// TIA Portal V19 export
// export: Created 2026-10-15T09:44:24.355296Z, ExportSetting WithDefaults, DisplayName Totally Integrated Automation Portal, DisplayVersion V19, DisplayName TIA Portal Openness, DisplayVersion V19, DisplayName TIA Portal Version Control Interface, DisplayVersion V19, DisplayName STEP 7 Professional, DisplayVersion V19, DisplayName STEP 7 Safety, DisplayVersion V19, DisplayName WinCC Basic/Comfort/Advanced, DisplayVersion V19, DisplayName WinCC Unified, DisplayVersion V19
FUNCTION "ROLL_PB16" : Void   // FC24, SCL
{ S7_Optimized_Access := 'TRUE' }
VERSION : 0.1
// stored: AutoNumber true, IsIECCheckEnabled false, SetENOAutomatically false, UDAEnableTagReadback false
   VAR_TEMP
      r : Bool;
      a1 : Word;
      a2 : Word;
      activeDataBlock : Int;
      comparisonResults : Array[0..0] of Bool;
   END_VAR
BEGIN

   #r := FALSE;
   #a1 := W#16#0000;
   #a2 := W#16#0000;
   #activeDataBlock := 0;
   // PB16, STEP 5 network 1
   #r := ("ROLL_IO".Input[0, 1] AND "ROLL_State".M[190, 5] AND "ROLL_State".M[190, 6] AND "ROLL_State".M[27, 7]);
   "ROLL_State".M[73, 7] := #r;
   // PB16, STEP 5 network 2
   #r := (("ROLL_State".M[20, 3] OR "ROLL_State".M[20, 5]) AND "ROLL_IO".Input[124, 1] AND "ROLL_IO".Input[124, 4]);
   "ROLL_State".M[74, 2] := #r;
   // PB16, STEP 5 network 3
   #r := (((NOT "ROLL_State".M[190, 5]) AND "ROLL_State".M[190, 6] AND "ROLL_State".M[74, 2]) OR (("ROLL_State".M[70, 2] OR "ROLL_State".M[70, 3]) AND "ROLL_State".M[74, 0]));
   "ROLL_State".M[74, 1] := #r;
   // PB16, STEP 5 network 4
   #r := (("ROLL_State".M[20, 4] OR "ROLL_State".M[20, 5]) AND "ROLL_IO".Input[0, 1] AND "ROLL_State".M[190, 6]);
   "ROLL_State".M[74, 4] := #r;
   // PB16, STEP 5 network 5
   #r := ((NOT "ROLL_IO".Output[113, 3]) AND ("ROLL_IO".Input[123, 6] OR "ROLL_State".M[70, 3] OR "ROLL_State".M[70, 5] OR "ROLL_State".M[70, 6]) AND ("ROLL_State".M[74, 0] OR "ROLL_State".M[74, 4]));
   "ROLL_State".M[74, 5] := #r;
   // PB16, STEP 5 network 6
   #r := ((NOT "ROLL_IO".Input[11, 0]) AND (NOT "ROLL_IO".Input[11, 1]) AND (NOT "ROLL_IO".Input[11, 2]) AND (NOT "ROLL_IO".Input[11, 3]) AND (NOT "ROLL_IO".Input[11, 4]) AND (NOT "ROLL_IO".Input[119, 6]) AND (NOT "ROLL_IO".Input[119, 7]) AND (NOT "ROLL_IO".Input[120, 0]) AND (NOT "ROLL_IO".Input[120, 1]));
   "ROLL_State".M[75, 2] := #r;
   // PB16, STEP 5 network 7
   #r := (("ROLL_State".M[190, 6] AND "ROLL_State".M[23, 1] AND "ROLL_State".M[75, 3]) OR "ROLL_State".M[75, 2]);
   "ROLL_State".M[75, 3] := #r;
   // PB16, STEP 5 network 8
   #r := ((((NOT "ROLL_IO".Input[11, 0]) AND (NOT "ROLL_IO".Input[11, 1]) AND (NOT "ROLL_IO".Input[11, 2]) AND (NOT "ROLL_IO".Input[11, 3]) AND (NOT "ROLL_IO".Input[11, 4]) AND (NOT "ROLL_IO".Input[119, 6]) AND (NOT "ROLL_IO".Input[119, 7]) AND (NOT "ROLL_IO".Input[120, 0]) AND (NOT "ROLL_IO".Input[120, 1]) AND "ROLL_IO".Input[13, 3]) OR "ROLL_State".M[63, 1]) AND ((NOT "ROLL_IO".Input[11, 6]) OR (NOT "ROLL_State".M[75, 3]) OR "ROLL_State".M[75, 2]) AND "ROLL_IO".Input[0, 1] AND "ROLL_IO".Input[12, 5] AND "ROLL_State".M[190, 6] AND "ROLL_State".M[23, 1]);
   "ROLL_State".M[75, 4] := #r;
   // PB16, STEP 5 network 9
   #r := ((((NOT "ROLL_IO".Input[11, 0]) AND (NOT "ROLL_IO".Input[11, 1]) AND (NOT "ROLL_IO".Input[11, 2]) AND (NOT "ROLL_IO".Input[11, 3]) AND (NOT "ROLL_IO".Input[11, 4]) AND (NOT "ROLL_IO".Input[119, 6]) AND (NOT "ROLL_IO".Input[119, 7]) AND (NOT "ROLL_IO".Input[120, 0]) AND (NOT "ROLL_IO".Input[120, 1]) AND "ROLL_IO".Input[13, 3]) OR "ROLL_State".M[63, 1]) AND (((NOT "ROLL_State".M[190, 6]) AND "ROLL_State".M[190, 5] AND "ROLL_State".M[23, 1]) OR "ROLL_State".M[74, 0]) AND "ROLL_IO".Input[0, 1]);
   "ROLL_State".M[75, 5] := #r;
   // PB16, STEP 5 network 10
   #r := (((NOT "ROLL_IO".Input[11, 0]) AND (("ROLL_IO".Input[0, 1] AND "ROLL_State".M[190, 5] AND "ROLL_State".M[23, 1]) OR "ROLL_State".M[74, 0]) AND "ROLL_State".M[63, 1]) OR ("ROLL_IO".Input[0, 1] AND "ROLL_State".M[190, 6] AND "ROLL_State".M[23, 1] AND "ROLL_State".M[75, 2]));
   "ROLL_State".M[75, 6] := #r;
   // PB16, STEP 5 network 11
   #r := ((NOT "ROLL_IO".Input[11, 0]) AND "ROLL_IO".Input[11, 6] AND "ROLL_State".M[190, 5] AND "ROLL_State".M[23, 0]);
   "ROLL_State".M[76, 0] := #r;
   // PB16, STEP 5 network 12
   #r := (((NOT "ROLL_IO".Input[11, 0]) AND "ROLL_State".M[74, 0]) OR ("ROLL_IO".Input[11, 0] AND "ROLL_IO".Input[11, 6] AND "ROLL_State".M[190, 6] AND "ROLL_State".M[23, 0]));
   "ROLL_State".M[76, 1] := #r;
   // PB16, STEP 5 network 13
   #r := (("ROLL_State".M[76, 0] OR "ROLL_State".M[76, 1]) AND "ROLL_IO".Input[0, 1]);
   "ROLL_State".M[76, 2] := #r;
   // PB16, STEP 5 network 14
   #r := ((NOT "ROLL_IO".Input[12, 1]) AND (NOT "ROLL_IO".Input[12, 5]));
   "ROLL_State".M[240, 0] := #r;
   // PB16, STEP 5 network 15
   #r := (("ROLL_State".M[190, 6] AND "ROLL_State".M[23, 0] AND "ROLL_State".M[77, 1]) OR "ROLL_State".M[240, 0]);
   "ROLL_State".M[77, 1] := #r;
   // PB16, STEP 5 network 16
   #r := ((((NOT "ROLL_IO".Input[12, 1]) AND ("ROLL_IO".Input[11, 1] OR "ROLL_IO".Input[11, 2] OR "ROLL_IO".Input[11, 3] OR "ROLL_IO".Input[11, 4] OR "ROLL_IO".Input[119, 6] OR "ROLL_IO".Input[119, 7] OR "ROLL_IO".Input[120, 0] OR "ROLL_IO".Input[120, 1])) OR (NOT "ROLL_IO".Input[12, 7])) AND ((NOT "ROLL_IO".Input[12, 7]) OR (NOT "ROLL_State".M[77, 1]) OR "ROLL_State".M[240, 0]) AND "ROLL_IO".Input[0, 1] AND "ROLL_IO".Input[11, 6] AND "ROLL_State".M[190, 6] AND "ROLL_State".M[23, 0]);
   "ROLL_State".M[77, 2] := #r;
   // PB16, STEP 5 network 17
   #r := (((NOT "ROLL_State".M[6, 0]) AND (NOT "ROLL_State".M[6, 2]) AND ("ROLL_IO".Input[11, 1] OR "ROLL_IO".Input[11, 2] OR "ROLL_IO".Input[11, 3] OR "ROLL_IO".Input[11, 4] OR "ROLL_IO".Input[119, 6] OR "ROLL_IO".Input[119, 7] OR "ROLL_IO".Input[120, 0])) OR "ROLL_IO".Input[11, 4]);
   "ROLL_State".M[76, 4] := #r;
   // PB16, STEP 5 network 18
   #r := ((NOT "ROLL_State".M[190, 5]) AND "ROLL_State".M[190, 6] AND "ROLL_State".M[23, 0] AND "ROLL_State".M[76, 4] AND "ROLL_State".M[77, 2]);
   "ROLL_State".M[76, 5] := #r;
   // PB16, STEP 5 network 19
   #r := ((((NOT "ROLL_State".M[190, 6]) AND "ROLL_State".M[190, 5] AND "ROLL_State".M[23, 0]) OR "ROLL_State".M[74, 0]) AND (("ROLL_IO".Input[124, 2] AND "ROLL_IO".Input[124, 5]) OR "ROLL_State".M[0, 4]) AND "ROLL_IO".Input[11, 0] AND "ROLL_State".M[63, 1]);
   "ROLL_State".M[76, 6] := #r;
   // PB16, STEP 5 network 20
   #r := (((((NOT "ROLL_IO".Input[12, 1]) OR (NOT "ROLL_IO".Input[12, 7])) AND "ROLL_State".M[76, 6]) OR "ROLL_State".M[76, 5]) AND "ROLL_IO".Input[0, 1] AND "ROLL_IO".Input[11, 6]);
   "ROLL_State".M[77, 0] := #r;
   // PB16, STEP 5 network 21
   #r := (((NOT "ROLL_IO".Input[11, 0]) AND (NOT "ROLL_IO".Input[12, 5]) AND "ROLL_State".M[190, 5]) OR ((NOT "ROLL_IO".Input[12, 1]) AND "ROLL_IO".Input[11, 0] AND "ROLL_State".M[190, 6]));
   "ROLL_State".M[240, 0] := #r;
   // PB16, STEP 5 network 22
   #r := ((NOT "ROLL_IO".Input[12, 1]) AND ("ROLL_IO".Input[11, 1] OR "ROLL_IO".Input[11, 2] OR "ROLL_IO".Input[11, 3] OR "ROLL_IO".Input[11, 4] OR "ROLL_IO".Input[119, 6] OR "ROLL_IO".Input[119, 7] OR "ROLL_IO".Input[120, 0]));
   "ROLL_State".M[240, 1] := #r;
   // PB16, STEP 5 network 23
   #r := ((NOT "ROLL_IO".Input[12, 1]) AND "ROLL_IO".Input[11, 0]);
   "ROLL_State".M[240, 2] := #r;
   // PB16, STEP 5 network 24
   #r := ((("ROLL_State".M[240, 1] OR "ROLL_State".M[240, 2]) AND "ROLL_State".M[77, 0]) OR ("ROLL_State".M[240, 0] AND "ROLL_State".M[76, 2]));
   "ROLL_State".M[76, 7] := #r;
   // PB16, STEP 5 network 25
   #r := ((NOT "ROLL_IO".Output[113, 3]) AND (NOT "ROLL_State".M[70, 2]) AND (NOT "ROLL_State".M[70, 3]) AND "ROLL_IO".Input[0, 1] AND "ROLL_IO".Input[11, 0] AND "ROLL_IO".Input[12, 1] AND "ROLL_IO".Input[12, 7] AND "ROLL_IO".Input[124, 5]);
   "ROLL_State".M[77, 3] := #r;
   // PB16, STEP 5 network 26
   #r := ((NOT "ROLL_State".M[77, 6]) AND (((NOT "ROLL_State".M[190, 6]) AND "ROLL_State".M[190, 5] AND "ROLL_State".M[22, 0]) OR "ROLL_State".M[74, 0]) AND "ROLL_IO".Output[113, 2] AND "ROLL_State".M[77, 3]);
   "ROLL_State".M[77, 4] := #r;
   // PB16, STEP 5 network 27
   #r := ((NOT "ROLL_State".M[190, 5]) AND (NOT "ROLL_State".M[77, 4]) AND "ROLL_State".M[190, 6] AND "ROLL_State".M[22, 0] AND "ROLL_State".M[77, 3]);
   "ROLL_State".M[77, 6] := #r;
   // PB16, STEP 5 network 28
   #r := ((NOT "ROLL_IO".Input[124, 5]) AND (NOT "ROLL_State".M[70, 3]) AND (((NOT "ROLL_IO".Input[124, 4]) AND "ROLL_State".M[20, 2] AND "ROLL_State".M[74, 0]) OR ((NOT "ROLL_State".M[190, 5]) AND "ROLL_IO".Input[0, 1] AND "ROLL_State".M[190, 6] AND "ROLL_State".M[22, 1])) AND "ROLL_IO".Input[124, 1]);
   "ROLL_State".M[77, 7] := #r;
   // PB16, STEP 5 network 29
   #r := ((NOT "ROLL_IO".Input[124, 4]) AND (NOT "ROLL_State".M[70, 3]) AND (((NOT "ROLL_State".M[15, 1]) AND "ROLL_State".M[20, 1] AND "ROLL_State".M[74, 0]) OR ((NOT "ROLL_State".M[190, 6]) AND "ROLL_IO".Input[0, 1] AND "ROLL_State".M[190, 5] AND "ROLL_State".M[22, 1])) AND "ROLL_IO".Input[124, 1]);
   "ROLL_State".M[78, 0] := #r;
   // PB16, STEP 5 network 30
   #r := ((("ROLL_State".M[22, 3] OR "ROLL_State".M[22, 4]) AND "ROLL_IO".Input[0, 1] AND "ROLL_State".M[190, 6]) OR ("ROLL_IO".Input[123, 5] AND "ROLL_State".M[74, 0]));
   IF #r THEN
       "ROLL_State".M[78, 4] := TRUE;
   END_IF;
   #r := (((NOT "ROLL_IO".Output[113, 3]) AND (NOT "ROLL_IO".Input[123, 4]) AND "ROLL_State".M[74, 0]) OR ((NOT "ROLL_IO".Output[113, 3]) AND "ROLL_IO".Input[0, 1] AND "ROLL_State".M[190, 5] AND "ROLL_State".M[22, 3]) OR (NOT "ROLL_IO".Input[0, 1]));
   IF #r THEN
       "ROLL_State".M[78, 4] := FALSE;
   END_IF;
   // PB16, STEP 5 network 31
   #r := ((NOT "ROLL_IO".Input[123, 5]) AND (NOT "ROLL_IO".Input[123, 6]) AND (NOT "ROLL_State".M[16, 0]) AND (NOT "ROLL_State".M[16, 4]) AND (NOT "ROLL_State".M[9, 1]) AND ((NOT "ROLL_IO".Input[123, 4]) OR "ROLL_State".M[190, 1]));
   "ROLL_State".M[78, 5] := #r;
   // PB16, STEP 5 network 32
   #r := (((NOT "ROLL_IO".Input[124, 2]) AND (NOT "ROLL_State".M[190, 5]) AND (NOT "ROLL_State".M[70, 3]) AND "ROLL_IO".Input[0, 1] AND "ROLL_IO".Input[124, 1] AND "ROLL_IO".Input[124, 4] AND "ROLL_State".M[190, 6] AND "ROLL_State".M[22, 4]) OR ("ROLL_State".M[70, 2] AND "ROLL_State".M[74, 0]));
   IF #r THEN
       "ROLL_State".M[78, 6] := TRUE;
   END_IF;
   #r := (((NOT "ROLL_State".M[70, 2]) AND ((NOT "ROLL_IO".Input[124, 1]) OR (NOT "ROLL_IO".Input[124, 4])) AND "ROLL_State".M[20, 2] AND "ROLL_State".M[74, 0]) OR ((NOT "ROLL_State".M[70, 2]) AND "ROLL_IO".Input[0, 1] AND "ROLL_State".M[190, 5] AND "ROLL_State".M[22, 4]) OR ((NOT "ROLL_State".M[70, 2]) AND "ROLL_State".M[20, 1] AND "ROLL_State".M[74, 0]) OR (NOT "ROLL_IO".Input[0, 1]) OR "ROLL_State".M[70, 0]);
   IF #r THEN
       "ROLL_State".M[78, 6] := FALSE;
   END_IF;
   // PB16, STEP 5 network 33
   #r := (((NOT "ROLL_State".M[70, 2]) AND (("ROLL_IO".Input[124, 5] AND "ROLL_State".M[20, 2]) OR "ROLL_State".M[20, 1]) AND "ROLL_State".M[74, 0]) OR ((NOT "ROLL_State".M[70, 2]) AND "ROLL_IO".Input[0, 1] AND "ROLL_State".M[190, 5] AND "ROLL_State".M[22, 4]));
   IF #r THEN
       "ROLL_State".M[78, 7] := TRUE;
   END_IF;
   #r := ((NOT "ROLL_IO".Input[0, 1]) OR "ROLL_State".M[70, 0] OR "ROLL_State".M[78, 6]);
   IF #r THEN
       "ROLL_State".M[78, 7] := FALSE;
   END_IF;
   // PB16, STEP 5 network 34
   RETURN;
END_FUNCTION
